Fanuc KAREL source: KD00029.KL

PROGRAM KD00029
%NOLOCKGROUP
VAR
  I: INTEGER
  J: INTEGER
  B: BOOLEAN
  R: REAL
  S: STRING[80]
BEGIN
  CONDITION[1]:
  WHEN CONTINUE DO
    I = 1
  ENDCONDITION
END KD00029
